(* IEC 61131-3 sources: JingjiangArm/moonboxpro_arm_8.4/Application/Application/任务列表/LogTask/粗采样保存, 7 files *)

(* ---- StRSampData.st ---- *)
(*@CES
Name=StRSampData
Type=Gvl
TypeGuid=2db5746d-d284-4425-9f7f-2663a34b0ebc
Guid=647225e6-5d7c-4765-8d74-e5faea58caf3
HasDeclaration=True
HasImplementation=False
*)
{DECLARATION}
TYPE StRSampData :
STRUCT
	abyRs_T1: ARRAY[1..4000] OF BYTE;(* T1粗采样 *)
	abyRs_T2: ARRAY[1..4000] OF BYTE;(* T2粗采样 *)
	byUnitNR: BYTE;(* 色组号 *)
	diVel: DINT;(* 速度*100.0 *)
	udiTskCycleNR: UDINT;(* 任务周期计数 *)
END_STRUCT
END_TYPE
{IMPLEMENTATION}

(* ---- StRSampFifo.st ---- *)
(*@CES
Name=StRSampFifo
Type=Gvl
TypeGuid=2db5746d-d284-4425-9f7f-2663a34b0ebc
Guid=e00882fe-97d1-4528-b28a-72dc94cf0559
HasDeclaration=True
HasImplementation=False
*)
{DECLARATION}
TYPE StRSampFifo :
STRUCT
	byIDX_Wr: BYTE;(* 取低3bits/正常操作一直累加就ok *)
	byIDX_Rd: BYTE;(* 取低3bits/正常操作一直累加就ok *)
	astStRSampData: ARRAY [0..7] OF StRSampData;
END_STRUCT
END_TYPE
{IMPLEMENTATION}

(* ---- StSampleDataForTest.st ---- *)
(*@CES
Name=StSampleDataForTest
Type=Gvl
TypeGuid=2db5746d-d284-4425-9f7f-2663a34b0ebc
Guid=737cf5e7-7729-43ac-8b0b-9f7abe5c616b
HasDeclaration=True
HasImplementation=False
*)
{DECLARATION}
TYPE StSampleDataForTest :
STRUCT
	byIdx		: BYTE;(* 索引/只取低3位/有效范围0~7 *)
	abyBuf_Rs	: ARRAY [0..7,1..8000] OF BYTE;(* 粗采样数据缓存 *)
	abyBuf_Fs	: ARRAY [0..7,1..8000] OF BYTE;(* 精采样数据缓存 *)
END_STRUCT
END_TYPE
{IMPLEMENTATION}

(* ---- KESAI_GTSD_TEST_SAMPLE_VERSION.st ---- *)
(*@CES
Name=KESAI_GTSD_TEST_SAMPLE_VERSION
Type=FunctionBlock
TypeGuid=6f9dac99-8de1-4efc-8465-68ac443b7d08
Guid=003f5c8f-60a7-4511-9628-a8eb072fa6d2
HasDeclaration=True
HasImplementation=True
*)
{DECLARATION}
FUNCTION KESAI_GTSD_TEST_SAMPLE_VERSION : STRING
VAR_INPUT
END_VAR
VAR
END_VAR

{IMPLEMENTATION}
KESAI_GTSD_TEST_SAMPLE_VERSION:= 'KESAI_GTSD_TEST_SAMPLE VERSION@2022.4.8.211617';

(* ---- KS_InstallMem_RS.st ---- *)
(*@CES
Name=KS_InstallMem_RS
Type=FunctionBlock
TypeGuid=6f9dac99-8de1-4efc-8465-68ac443b7d08
Guid=3c1006dd-3441-469c-8106-999143937635
HasDeclaration=True
HasImplementation=True
*)
{DECLARATION}
FUNCTION KS_InstallMem_RS : INT
VAR_INPUT
	i_ppstStRSampFifo: POINTER TO POINTER TO StRSampFifo;
END_VAR
VAR
	iResult: INT;
	pstStRSampFifo_Tmp: POINTER TO StRSampFifo;
END_VAR
{IMPLEMENTATION}
IF i_ppstStRSampFifo<>0 THEN
	pstStRSampFifo_Tmp:= SysMemAlloc(SIZEOF(pstStRSampFifo_Tmp^));
	IF pstStRSampFifo_Tmp<>0 THEN
		pstStRSampFifo_Tmp^.byIDX_Wr:= 0;
		pstStRSampFifo_Tmp^.byIDX_Rd:= 0;
		i_ppstStRSampFifo^:= pstStRSampFifo_Tmp;
		iResult:= 0;
	ELSE
		iResult:= -2;(* 内存申请失败 *)
	END_IF
ELSE
	iResult:= -1;
END_IF
KS_InstallMem_RS:= iResult;

(* ---- KS_PshRSdata2Fifo.st ---- *)
(*@CES
Name=KS_PshRSdata2Fifo
Type=FunctionBlock
TypeGuid=6f9dac99-8de1-4efc-8465-68ac443b7d08
Guid=7d186a17-b9d1-422c-94b2-454e470a5b16
HasDeclaration=True
HasImplementation=True
*)
{DECLARATION}
FUNCTION KS_PshRSdata2Fifo : INT
VAR_INPUT
	i_pstStRSampFifo: POINTER TO StRSampFifo;
	i_pbyRs_T1: POINTER TO BYTE;
	i_pbyRs_T2: POINTER TO BYTE;
	i_byUnitNR: BYTE;
	i_diVel: DINT;
	i_udiTskCycleNR: UDINT;
END_VAR
VAR
	iResult: INT;
	byIDX_Tmp: BYTE;
END_VAR
{IMPLEMENTATION}
IF i_pstStRSampFifo<>0 AND
	i_pbyRs_T1<>0 AND
	i_pbyRs_T2<>0 THEN

	byIDX_Tmp:= i_pstStRSampFifo^.byIDX_Wr AND BYTE#7;(* 控制循环0~7 *)
	i_pstStRSampFifo^.astStRSampData[byIDX_Tmp].byUnitNR:= i_byUnitNR;
	i_pstStRSampFifo^.astStRSampData[byIDX_Tmp].diVel:= i_diVel;
	i_pstStRSampFifo^.astStRSampData[byIDX_Tmp].udiTskCycleNR:= i_udiTskCycleNR;
	SysMemCpy(
		ADR(i_pstStRSampFifo^.astStRSampData[byIDX_Tmp].abyRs_T1),
		i_pbyRs_T1,
		SIZEOF(i_pstStRSampFifo^.astStRSampData[byIDX_Tmp].abyRs_T1) );
	SysMemCpy(
		ADR(i_pstStRSampFifo^.astStRSampData[byIDX_Tmp].abyRs_T2),
		i_pbyRs_T2,
		SIZEOF(i_pstStRSampFifo^.astStRSampData[byIDX_Tmp].abyRs_T2) );

	i_pstStRSampFifo^.byIDX_Wr:= byIDX_Tmp+1;

	iResult:= 0;
ELSE
	iResult:= -1;
END_IF
KS_PshRSdata2Fifo:= iResult;

(* ---- KS_FB_ExportRSFifo2File.st ---- *)
(*@CES
Name=KS_FB_ExportRSFifo2File
Type=FunctionBlock
TypeGuid=6f9dac99-8de1-4efc-8465-68ac443b7d08
Guid=280a4f81-a5dc-40a5-adea-619cfced529e
HasDeclaration=True
HasImplementation=True
*)
{DECLARATION}
FUNCTION_BLOCK KS_FB_ExportRSFifo2File
VAR_INPUT
	i_xEn: BOOL;
	i_sPath: STRING :=  '/data/kesai/data/RS';
	i_pstStRSampFifo: POINTER TO StRSampFifo := 0;
END_VAR
VAR_OUTPUT
	//o_xEno: BOOL;
	o_iErNo: INT;(* 0表示ok/-1参数错误/-2文件创建失败/100暂时没有数据写入 *)
END_VAR
VAR
	byIDX_Wr_Tmp: BYTE;
	byIDX_Rd_Tmp: BYTE;
	sFullFname: STRING(260):= '';
	dwHdlFile: RTS_IEC_HANDLE;(* TYPE RTS_IEC_HANDLE : POINTER TO BYTE *)
	udiRtn: RTS_IEC_RESULT;(* TYPE RTS_IEC_RESULT : UDINT *)
						(* TYPE RTS_IEC_SIZE : POINTER TO BYTE *)
						(* RTS_INVALID_HANDLE: RTS_IEC_HANDLE(-1) *)
END_VAR
{IMPLEMENTATION}
IF i_xEn THEN
	IF i_pstStRSampFifo<>0 THEN
		byIDX_Wr_Tmp:= i_pstStRSampFifo^.byIDX_Wr AND BYTE#7;
		byIDX_Rd_Tmp:= i_pstStRSampFifo^.byIDX_Rd AND BYTE#7;
		IF byIDX_Wr_Tmp<>byIDX_Rd_Tmp THEN

			sFullFname:= i_sPath;
			IF RIGHT(i_sPath,1)<>'\' THEN
				sFullFname:= CONCAT(sFullFname, '\');
			END_IF
			sFullFname:= CONCAT(sFullFname, 'U');
			sFullFname:= CONCAT(sFullFname, BYTE_TO_STRING(i_pstStRSampFifo^.astStRSampData[byIDX_Rd_Tmp].byUnitNR));
			sFullFname:= CONCAT(sFullFname, '-');
			sFullFname:= CONCAT(sFullFname, UDINT_TO_STRING(i_pstStRSampFifo^.astStRSampData[byIDX_Rd_Tmp].udiTskCycleNR));
			sFullFname:= CONCAT(sFullFname, '-');
			sFullFname:= CONCAT(sFullFname, DINT_TO_STRING(i_pstStRSampFifo^.astStRSampData[byIDX_Rd_Tmp].diVel));
			sFullFname:= CONCAT(sFullFname, '@');
			sFullFname:= CONCAT(sFullFname, KS_GetTimeString(TIMEFORMAT_HYPHEN_DOT, TRUE, TRUE));
			sFullFname:= CONCAT(sFullFname, '.rs');

			dwHdlFile:= SysFileOpen(sFullFname, SysFile.AM_WRITE, ADR(udiRtn));
			IF dwHdlFile<>0 THEN
				SysFileWrite(
					dwHdlFile,
					ADR(i_pstStRSampFifo^.astStRSampData[byIDX_Rd_Tmp].abyRs_T1),
					SIZEOF(i_pstStRSampFifo^.astStRSampData[byIDX_Rd_Tmp].abyRs_T1),
					 ADR(udiRtn));
				SysFileWrite(
					dwHdlFile,
					ADR(i_pstStRSampFifo^.astStRSampData[byIDX_Rd_Tmp].abyRs_T2),
					SIZEOF(i_pstStRSampFifo^.astStRSampData[byIDX_Rd_Tmp].abyRs_T2),
					 ADR(udiRtn));
				SysFileClose(dwHdlFile);

				i_pstStRSampFifo^.byIDX_Rd:= byIDX_Rd_Tmp+1;
			ELSE
				o_iErNo:= -2;
			END_IF
		ELSE
			o_iErNo:= 100;
		END_IF
	ELSE
		o_iErNo:= -1;
	END_IF
END_IF
